PROGRAM MAIN
VAR
END_VAR

PRG_Echo();
PRG_EchoMqtt();

END_PROGRAM

(* stored: Version 1.1.0.1
   POU MAIN: Id {5f84cfb4-87d6-48cc-aa81-ab9446558539}, SpecialFunc None *)
